// FB_Hrl - the whole practice plant as the root mode node: one aisle with one
// RBG, the rack, the pre-zone with I-point and in-feed/out-feed conveyors, and
// the MFR interface.
// Pre-zone flow: in-feed (pallet already checked at the I-point) -> transfer
// station -> RBG stores it. Retrieved pallets are put on the station and leave
// over the out-feed.
FUNCTION_BLOCK FB_Hrl EXTENDS FB_ModeNode
VAR_INPUT
    stConfig : ST_HrlConfig;   // applied once on the first cycle (set it before)
    sConfigError : STRING(120);   // from FB_HrlConfig; shown as a fault
    stSafety     : ST_SafetyStatus;   // map from the safety controller (TwinSAFE group outputs)
    bSafetyReset : BOOL;              // acknowledge button
    bDoorRequest : BOOL;              // operator wants to enter the aisle
END_VAR
VAR
    fbRack    : FB_Rack;
    fbSrm     : FB_Srm(ipParent := THIS^, sNodeName := 'RBG01');
    fbInfeed  : FB_ConveyorZone(ipParent := THIS^, sNodeName := 'Infeed');
    fbOutfeed : FB_ConveyorZone(ipParent := THIS^, sNodeName := 'Outfeed');
    fbIPoint  : FB_IPoint;
    fbMfr     : FB_MfrInterface;
    fbMfrTcp  : FB_MfrLinkTcp;     // used when stConfig.eMfrLink = eTcp
    fbTeach   : FB_TeachIn;        // guided teach-in (manual mode)
    fbDiag    : FB_Diag;           // active faults for the HMI + TwinCAT logger
    fbSafety  : FB_SafetyInterface;
    bInitDone : BOOL;
    nInStep   : INT;
    sMovingLe : STRING(20);
END_VAR
VAR_OUTPUT
    bStationOutbound : BOOL;   // pallet on the station is leaving (retrieved), not arriving
    bStationReserved : BOOL;   // station held free for a retrieval: the in-feed must wait
    bSafetyOk        : BOOL;   // drives may run; FALSE -> MAIN forces stop mode
    bDoorUnlockReq   : BOOL;   // to the safety controller
END_VAR

METHOD PROTECTED OnCyclic
VAR_INPUT
END_VAR
IF NOT bInitDone THEN
    // The plant is built from the configuration; the code below never changes per site.
    fbRack.stCfg      := stConfig.stRack;
    fbSrm.eAxisKind   := stConfig.eAxisKind;
    fbSrm.stTravelCfg := stConfig.stTravel;
    fbSrm.stHoistCfg  := stConfig.stHoist;
    fbSrm.stForkCfg   := stConfig.stFork;
    ApplyZone(fbInfeed, stConfig.stInfeed);    // same standard block, other parameters
    ApplyZone(fbOutfeed, stConfig.stOutfeed);
    fbMfr.lrAckTimeout := stConfig.lrAckTimeout;
    fbSrm.Init(fbRack);
    fbMfr.Init(fbRack, fbSrm);
    fbTeach.Init(fbRack, fbSrm);
    fbMfrTcp.nPort    := stConfig.nMfrPort;
    fbMfrTcp.stLayout := stConfig.stLayout;
    bInitDone := TRUE;
END_IF
IF stConfig.eMfrLink = E_MfrLink.eTcp THEN
    fbMfrTcp.Cyclic();          // the link stays up in every operating mode
    fbMfr.Serve(fbMfrTcp);
END_IF
fbSafety(stStatus := stSafety, bSimulate := stConfig.bSafetySimulate, bReset := bSafetyReset,
         bDoorRequest := bDoorRequest, bStandstill := NOT fbSrm.bBusy AND NOT fbSrm.bGotoActive);
bSafetyOk      := fbSafety.bDriveEnable;
bDoorUnlockReq := fbSafety.bDoorUnlockReq;
SUPER^.OnCyclic();
fbDiag.Check(E_Fault.eSafety, NOT bSafetyOk, 'Safety stop - check e-stop and aisle door, then acknowledge');
fbDiag.Check(E_Fault.eSrmAxis, fbSrm.bFault, 'RBG axis fault - check the drive, then ResetFault');
fbDiag.Check(E_Fault.eInfeedJam, fbInfeed.eState = E_ZoneState.eFault, 'In-feed jam - clear the pallet, reset the zone');
fbDiag.Check(E_Fault.eOutfeedJam, fbOutfeed.eState = E_ZoneState.eFault, 'Out-feed jam - clear the pallet, reset the zone');
fbDiag.Check(E_Fault.eMfrAck, fbMfr.bAckTimeout, 'MFR did not acknowledge TDON - check the MFR');
fbDiag.Check(E_Fault.eMfrLinkDown, stConfig.eMfrLink = E_MfrLink.eTcp AND NOT fbMfrTcp.bConnected,
             'No MFR connected - check network / MFR port');
fbDiag.Check(E_Fault.eConfig, sConfigError <> '', 'HrlConfig.json rejected - defaults in use, see sConfigError');
fbDiag.Check(E_Fault.eTeachRejected, fbTeach.bLastRejected, 'Teach-in refused - place too far from drawing, check rack');
END_METHOD

METHOD PROTECTED RunAutomatic
VAR_INPUT
END_VAR
VAR
    stStation : ST_SlotAddr := (nSide := 1, nColumn := 0, nLevel := 1);
END_VAR
fbMfr.Cyclic();

// In-feed -> transfer station
CASE nInStep OF
    0:  IF fbInfeed.eState = E_ZoneState.eOccupied AND NOT fbRack.IsOccupied(stStation)
           AND NOT bStationOutbound AND NOT bStationReserved THEN
            sMovingLe := fbInfeed.sLeId;
            nInStep   := 1;
        END_IF
    // Done once our pallet has left the zone. The previous zone may hand over
    // the next pallet in the same cycle, so "zone empty" alone can be missed.
    1:  IF fbInfeed.Deliver() = E_CmdResult.eDone OR fbInfeed.sLeId <> sMovingLe THEN
            fbRack.Put(stStation, sMovingLe);
            nInStep := 0;
        END_IF
END_CASE

// Transfer station -> out-feed (only pallets the RBG brought out)
IF bStationOutbound AND fbRack.IsOccupied(stStation)
   AND fbOutfeed.eState = E_ZoneState.eEmpty THEN
    fbOutfeed.Accept(fbRack.Take(stStation));
    bStationOutbound := FALSE;
    bStationReserved := FALSE;   // station free for the in-feed again
END_IF
IF fbOutfeed.eState = E_ZoneState.eOccupied THEN
    fbOutfeed.Deliver();   // goods-out takes it away
END_IF
END_METHOD

// Called when a retrieval to the station is ordered: that pallet leaves.
METHOD PUBLIC MarkStationOutbound
VAR_INPUT
END_VAR
bStationOutbound := TRUE;
END_METHOD

// Hold the transfer station free for the next retrieval. Without this the
// in-feed refills the station every time the RBG picks a pallet from it, and
// a retrieval never finds the station empty.
METHOD PUBLIC ReserveStation
VAR_INPUT
END_VAR
bStationReserved := TRUE;
END_METHOD

// Manual jog request from the HMI (acts in manual mode only).
METHOD PUBLIC Jog
VAR_INPUT
    eAxis : E_JogAxis;
    bFwd  : BOOL;
    bBwd  : BOOL;
END_VAR
fbSrm.eJogAxis := eAxis;
fbSrm.bJogFwd  := bFwd;
fbSrm.bJogBwd  := bBwd;
END_METHOD

METHOD PRIVATE ApplyZone
VAR_IN_OUT
    fbZone : FB_ConveyorZone;
END_VAR
VAR_INPUT
    stCfg : ST_ZoneConfig;
END_VAR
fbZone.lrLength     := stCfg.lrLength;
fbZone.lrSpeed      := stCfg.lrSpeed;
fbZone.lrJamTimeout := stCfg.lrJamTimeout;
fbZone.bSimulate    := stCfg.bSimulate;
END_METHOD

END_FUNCTION_BLOCK

(* stored: Version 1.1.0.1
   POU FB_Hrl: Id {8b101ed3-d0e1-44fa-8906-694294c7c611}, SpecialFunc None
   Method OnCyclic: Id {6e601098-e9b4-4401-8f54-1716c269968e}
   Method RunAutomatic: Id {10d74ef1-ca39-4c08-9fa9-d5ebb774ba3d}
   Method MarkStationOutbound: Id {88a3f4f0-41da-44c6-9d25-202279366aa0}
   Method ReserveStation: Id {3c1f6a52-8e0d-4b7a-9f31-5d2e7a90c4b8}
   Method Jog: Id {f83f1014-3638-d543-7b69-b77a7040e8d1}
   Method ApplyZone: Id {d2acfcce-701a-a281-639c-c14150369c7e} *)
